(* IEC 61131-3 sources: codesys-to-astra/tools/tests/fixtures/lowering/src/POUs/F_Noop, 1 file *)

(* ---- F_Noop.decl.st ---- *)
// Назначение: пример для понижения iec-checker (tools/tests/test_assemble.py)
// Автор:      kr0nsch
// Версия:     0.1.0
// Документ:   docs/LAYOUT.md, раздел «Собранный текст build/assembled»; tools/README.md
FUNCTION F_Noop : BOOL
VAR_INPUT
    xIn : BOOL;
END_VAR
